TYPE ET_BECKHOFF_AxisGetLimits :
(
	eWaitExecute := 0,
	eReadVeloMax,
	eWfReadVeloMax,
	eReadAccMax,
	eWfReadAccMax,
	eReadDecMax,
	eWfReadDecMax,
	eReadJerkMax,
	eWfReadJerkMax,
	eReadSoftLimitMax,
	eWfReadSoftLimitMax,
	eReadSoftLimitMin,
	eWfReadSoftLimitMin,
	eDone := 197,
	eError := 198,
	eNoExecute := 199
);
END_TYPE

(* stored: Version 1.1.0.1, ProductVersion 3.1.4024.15
   DUT ET_BECKHOFF_AxisGetLimits: Id {b7bfaed4-09d5-4532-8c3c-4e538f18a63a} *)
